// TIA Portal V14 SP1 export
// export: Created 2000-01-01T00:00:00.0000000Z, ExportSetting None
FUNCTION "FC_Rung" : Void   // FC42, LAD
{ S7_Optimized_Access := 'TRUE' }
   VAR_INPUT
      Local : Int;
   END_VAR
BEGIN

REGION Network 1
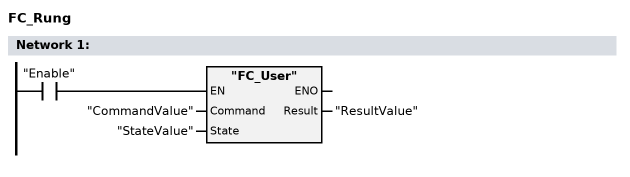
   RUNG wire#powerrail
      Contact( "Enable" )
      "FC_User"(Command := "CommandValue", State := "StateValue", Result => "ResultValue")
   END_RUNG
   // the same network as SCL:
   IF "Enable" THEN
       "FC_User"(Command := "CommandValue", State := "StateValue", Result => "ResultValue");
   END_IF;
END_REGION
END_FUNCTION
